Fanuc KAREL source: KT00434.KL

PROGRAM KT00434
%NOLOCKGROUP
VAR
  P1: JOINTPOS
  P2: JOINTPOS
  OUT: BOOLEAN
BEGIN
  OUT = P1 > P2
END KT00434
